Fanuc KAREL source: KA00198.KL

PROGRAM KA00198
%NOLOCKGROUP
VAR
  SRC: ARRAY[4] OF SHORT
  DST: ARRAY[4] OF JOINTPOS
BEGIN
  DST = SRC
END KA00198
